ABB RAPID module: Count_only_movec.mod

%%%
  VERSION:1
  LANGUAGE:ENGLISH
%%%
MODULE MOD_Count_only_movec

    ! -------------------------------
    ! Define customized variables here
    ! ...

	! Tool variables:

	! Reference variables:

	PROC Main()
		ConfJ \On;
		ConfL \Off;
		! Program generated by RoboDK v6.0.7 for ABB IRB 120-3/0.6 on XX/XX/XXXX 12:58:43
		! Using nominal kinematics.
		MoveC [[-618.417,609.652,333.231],[0.40821789,0.23456972,0.87542610,-0.10938165],[0,-1,0,0],[9E+09,9E+09,9E+09,9E+09,9E+09,9E+09]],[[-671.251,582.420,294.929],[0.40821789,0.23456972,0.87542610,-0.10938165],[0,-1,0,0],[9E+09,9E+09,9E+09,9E+09,9E+09,9E+09]],v500,z1,tool0 \WObj:=wobj0;
	ENDPROC

ENDMODULE
